(* IEC 61131-3 sources: SRCI_CLIENT_PLC/RobotLibrary/Library/Structures/Common, 4 files *)

(* ---- CmdHeader.st ---- *)
{attribute 'pack_mode' := '1'}
// -------------------------------------------------------------------------
//  SRCI Robot Library
// -------------------------------------------------------------------------
//
//  Object:      CmdHeader
//  Author:      Thorsten Brach
//  Date:        2024-06-01
//
//  Description:
//
//
//  Copyright:
//    (C) 2024 Thorsten Brach. All rights reserved
//             Licensed under the MIT License.
//
//  Disclaimer:
//    This project is provided without any guarantee and can be used for
//    private and commercial purposes. Any use is at the user’s
//    own risk and responsibility.
//
// -------------------------------------------------------------------------
TYPE CmdHeader :
STRUCT
  /// Type of command - For more information see chapter 5.6.4.
 CmdTyp          : CmdType;
 /// Specifies target buffer and processing behavior - For more information see chapter 5.6.4.5
 ExecMode        : ExecutionMode;
 /// Parameter Sequence, used to identify sets of CMD parameter
 ParSeq          : BYTE;
 /// Priority of this command
 Priority        : PriorityLevel;
END_STRUCT
END_TYPE

(* ---- LogParameter.st ---- *)
{attribute 'pack_mode' := '1'}
// -------------------------------------------------------------------------
//  SRCI Robot Library
// -------------------------------------------------------------------------
//
//  Object:      LogParameter
//  Author:      Thorsten Brach
//  Date:        2024-06-01
//
//  Description:
//
//
//  Copyright:
//    (C) 2024 Thorsten Brach. All rights reserved
//             Licensed under the MIT License.
//
//  Disclaimer:
//    This project is provided without any guarantee and can be used for
//    private and commercial purposes. Any use is at the user’s
//    own risk and responsibility.
//
// -------------------------------------------------------------------------
TYPE LogParameter :
STRUCT
  /// Log level setting for creating commands
  CreateCmd : LogLevel;
  /// Log level setting for updating commands
  UpdateCmd : LogLevel;
  /// Log level setting for generating sequence
  GenSeq    : LogLevel;
  /// Log level for ??? sequence
  DecSeq    : LogLevel;
END_STRUCT
END_TYPE

(* ---- RobotCoordinateSystemParameters.st ---- *)
{attribute 'pack_mode' := '1'}
// -------------------------------------------------------------------------
//  SRCI Robot Library
// -------------------------------------------------------------------------
//
//  Object:      RobotCoordinateSystemParameters
//  Author:      Thorsten Brach
//  Date:        2024-06-01
//
//  Description:
//
//
//  Copyright:
//    (C) 2024 Thorsten Brach. All rights reserved
//             Licensed under the MIT License.
//
//  Disclaimer:
//    This project is provided without any guarantee and can be used for
//    private and commercial purposes. Any use is at the user’s
//    own risk and responsibility.
//
// -------------------------------------------------------------------------
TYPE RobotCoordinateSystemParameters :
STRUCT
  /// Index of target tool
  /// • 0: Flange (default)
  /// • 1..254: Tool frames
  ToolNo : USINT;
  /// Index of target frame
  /// • 0: WCS (default)
  /// • 1..254: User frames
  FrameNo : USINT;
END_STRUCT
END_TYPE

(* ---- RspHeader.st ---- *)
{attribute 'pack_mode' := '1'}
// -------------------------------------------------------------------------
//  SRCI Robot Library
// -------------------------------------------------------------------------
//
//  Object:      RspHeader
//  Author:      Thorsten Brach
//  Date:        2024-06-01
//
//  Description:
//
//
//  Copyright:
//    (C) 2024 Thorsten Brach. All rights reserved
//             Licensed under the MIT License.
//
//  Disclaimer:
//    This project is provided without any guarantee and can be used for
//    private and commercial purposes. Any use is at the user’s
//    own risk and responsibility.
//
// -------------------------------------------------------------------------
TYPE RspHeader :
STRUCT
  /// Parameter Sequence, used to identify sets of CMD parameter - For more information see chapter 5.6.4
  ParSeq               : USINT;
  /// Actual state of the command - For more information and examples, see chapter 5.6.4.3
  State                : CmdMessageState;
  /// Severity of returned message according to .Table 5-49.
  AlarmMessageSeverity : Severity;
  /// Message code for error/warning/info identification reported during execution of command according to
  /// • Error: Table 7-1
  /// • Warning: Table 7-3
  /// • Info: Table 7-5
  AlarmMessageCode     : UINT;
END_STRUCT
END_TYPE
